{attribute 'qualified_only'}
{attribute 'strict'}
{attribute 'to_string'}
TYPE XtsHardwareDiscoveryState :
(
	WaitingForXpu := 0,
	GettingParts := 1,
	InitialisingXtsParts := 2,
	GettingTracks := 3,
	InitialisingXtsTracks := 4,
	GettingModules := 5,
	InitialisingModules := 6,
	GettingMovers := 7,
	InitialisingMovers := 8,	
	HardwareFound := 9,
	DiscoveryFault := 99,
	DiscoveryFailed := 999
);
END_TYPE

(* stored: Version 1.1.0.1
   DUT XtsHardwareDiscoveryState: Id {7cad66c2-2e7c-408e-8aec-b9645f1a57db} *)
